TYPE "UDT_Service_ControlBlockMedium"
VERSION : 0.1
   STRUCT
      mode : Int := 1;   //  Service/Mapping selection
      stepOrder { S7_SetPoint := 'False'} : "UDT_Service_StepOrderRawDataMedium";   // Configuration step order
      step { S7_SetPoint := 'False'} : "UDT_Service_StepRawDataMedium" := ([([16#FFFFFFFF], [16#FFFFFFFF], [16#FFFFFFFF], [16#FFFFFFFF]), ([16#FFFFFFFF], [16#FFFFFFFF], [16#FFFFFFFF], [16#FFFFFFFF]), ([16#FFFFFFFF], [16#FFFFFFFF], [16#FFFFFFFF], [16#FFFFFFFF]), ([16#FFFFFFFF], [16#FFFFFFFF], [16#FFFFFFFF], [16#FFFFFFFF]), ([16#FFFFFFFF], [16#FFFFFFFF], [16#FFFFFFFF], [16#FFFFFFFF]), ([16#FFFFFFFF], [16#FFFFFFFF], [16#FFFFFFFF], [16#FFFFFFFF]), ([16#FFFFFFFF], [16#FFFFFFFF], [16#FFFFFFFF], [16#FFFFFFFF]), ([16#FFFFFFFF], [16#FFFFFFFF], [16#FFFFFFFF], [16#FFFFFFFF]), ([16#FFFFFFFF], [16#FFFFFFFF], [16#FFFFFFFF], [16#FFFFFFFF]), ([16#FFFFFFFF], [16#FFFFFFFF], [16#FFFFFFFF], [16#FFFFFFFF]), ([16#FFFFFFFF], [16#FFFFFFFF], [16#FFFFFFFF], [16#FFFFFFFF]), ([16#FFFFFFFF], [16#FFFFFFFF], [16#FFFFFFFF], [16#FFFFFFFF]), ([16#FFFFFFFF], [16#FFFFFFFF], [16#FFFFFFFF], [16#FFFFFFFF]), ([16#FFFFFFFF], [16#FFFFFFFF], [16#FFFFFFFF], [16#FFFFFFFF]), ([16#FFFFFFFF], [16#FFFFFFFF], [16#FFFFFFFF], [16#FFFFFFFF]), ([16#FFFFFFFF], [16#FFFFFFFF], [16#FFFFFFFF], [16#FFFFFFFF]), ([16#FFFFFFFF], [16#FFFFFFFF], [16#FFFFFFFF], [16#FFFFFFFF]), ([16#FFFFFFFF], [16#FFFFFFFF], [16#FFFFFFFF], [16#FFFFFFFF]), ([16#FFFFFFFF], [16#FFFFFFFF], [16#FFFFFFFF], [16#FFFFFFFF]), ([16#FFFFFFFF], [16#FFFFFFFF], [16#FFFFFFFF], [16#FFFFFFFF]), ([16#FFFFFFFF], [16#FFFFFFFF], [16#FFFFFFFF], [16#FFFFFFFF]), ([16#FFFFFFFF], [16#FFFFFFFF], [16#FFFFFFFF], [16#FFFFFFFF]), ([16#FFFFFFFF], [16#FFFFFFFF], [16#FFFFFFFF], [16#FFFFFFFF]), ([16#FFFFFFFF], [16#FFFFFFFF], [16#FFFFFFFF], [16#FFFFFFFF]), ([16#FFFFFFFF], [16#FFFFFFFF], [16#FFFFFFFF], [16#FFFFFFFF]), ([16#FFFFFFFF], [16#FFFFFFFF], [16#FFFFFFFF], [16#FFFFFFFF]), ([16#FFFFFFFF], [16#FFFFFFFF], [16#FFFFFFFF], [16#FFFFFFFF]), ([16#FFFFFFFF], [16#FFFFFFFF], [16#FFFFFFFF], [16#FFFFFFFF]), ([16#FFFFFFFF], [16#FFFFFFFF], [16#FFFFFFFF], [16#FFFFFFFF]), ([16#FFFFFFFF], [16#FFFFFFFF], [16#FFFFFFFF], [16#FFFFFFFF]), ([16#FFFFFFFF], [16#FFFFFFFF], [16#FFFFFFFF], [16#FFFFFFFF]), ([16#FFFFFFFF], [16#FFFFFFFF], [16#FFFFFFFF], [16#FFFFFFFF]), ([16#FFFFFFFF], [16#FFFFFFFF], [16#FFFFFFFF], [16#FFFFFFFF]), ([16#FFFFFFFF], [16#FFFFFFFF], [16#FFFFFFFF], [16#FFFFFFFF]), ([16#FFFFFFFF], [16#FFFFFFFF], [16#FFFFFFFF], [16#FFFFFFFF]), ([16#FFFFFFFF], [16#FFFFFFFF], [16#FFFFFFFF], [16#FFFFFFFF]), ([16#FFFFFFFF], [16#FFFFFFFF], [16#FFFFFFFF], [16#FFFFFFFF]), ([16#FFFFFFFF], [16#FFFFFFFF], [16#FFFFFFFF], [16#FFFFFFFF]), ([16#FFFFFFFF], [16#FFFFFFFF], [16#FFFFFFFF], [16#FFFFFFFF]), ([16#FFFFFFFF], [16#FFFFFFFF], [16#FFFFFFFF], [16#FFFFFFFF]), ([16#FFFFFFFF], [16#FFFFFFFF], [16#FFFFFFFF], [16#FFFFFFFF]), ([16#FFFFFFFF], [16#FFFFFFFF], [16#FFFFFFFF], [16#FFFFFFFF]), ([16#FFFFFFFF], [16#FFFFFFFF], [16#FFFFFFFF], [16#FFFFFFFF]), ([16#FFFFFFFF], [16#FFFFFFFF], [16#FFFFFFFF], [16#FFFFFFFF]), ([16#FFFFFFFF], [16#FFFFFFFF], [16#FFFFFFFF], [16#FFFFFFFF]), ([16#FFFFFFFF], [16#FFFFFFFF], [16#FFFFFFFF], [16#FFFFFFFF]), ([16#FFFFFFFF], [16#FFFFFFFF], [16#FFFFFFFF], [16#FFFFFFFF]), ([16#FFFFFFFF], [16#FFFFFFFF], [16#FFFFFFFF], [16#FFFFFFFF]), ([16#FFFFFFFF], [16#FFFFFFFF], [16#FFFFFFFF], [16#FFFFFFFF]), ([16#FFFFFFFF], [16#FFFFFFFF], [16#FFFFFFFF], [16#FFFFFFFF]), ([16#FFFFFFFF], [16#FFFFFFFF], [16#FFFFFFFF], [16#FFFFFFFF]), ([16#FFFFFFFF], [16#FFFFFFFF], [16#FFFFFFFF], [16#FFFFFFFF]), ([16#FFFFFFFF], [16#FFFFFFFF], [16#FFFFFFFF], [16#FFFFFFFF]), ([16#FFFFFFFF], [16#FFFFFFFF], [16#FFFFFFFF], [16#FFFFFFFF]), ([16#FFFFFFFF], [16#FFFFFFFF], [16#FFFFFFFF], [16#FFFFFFFF]), ([16#FFFFFFFF], [16#FFFFFFFF], [16#FFFFFFFF], [16#FFFFFFFF]), ([16#FFFFFFFF], [16#FFFFFFFF], [16#FFFFFFFF], [16#FFFFFFFF]), ([16#FFFFFFFF], [16#FFFFFFFF], [16#FFFFFFFF], [16#FFFFFFFF]), ([16#FFFFFFFF], [16#FFFFFFFF], [16#FFFFFFFF], [16#FFFFFFFF]), ([16#FFFFFFFF], [16#FFFFFFFF], [16#FFFFFFFF], [16#FFFFFFFF]), ([16#FFFFFFFF], [16#FFFFFFFF], [16#FFFFFFFF], [16#FFFFFFFF]), ([16#FFFFFFFF], [16#FFFFFFFF], [16#FFFFFFFF], [16#FFFFFFFF]), ([16#FFFFFFFF], [16#FFFFFFFF], [16#FFFFFFFF], [16#FFFFFFFF]), ([16#FFFFFFFF], [16#FFFFFFFF], [16#FFFFFFFF], [16#FFFFFFFF]), ([16#FFFFFFFF], [16#FFFFFFFF], [16#FFFFFFFF], [16#FFFFFFFF]), ([16#FFFFFFFF], [16#FFFFFFFF], [16#FFFFFFFF], [16#FFFFFFFF]), ([16#FFFFFFFF], [16#FFFFFFFF], [16#FFFFFFFF], [16#FFFFFFFF]), ([16#FFFFFFFF], [16#FFFFFFFF], [16#FFFFFFFF], [16#FFFFFFFF]), ([16#FFFFFFFF], [16#FFFFFFFF], [16#FFFFFFFF], [16#FFFFFFFF]), ([16#FFFFFFFF], [16#FFFFFFFF], [16#FFFFFFFF], [16#FFFFFFFF]), ([16#FFFFFFFF], [16#FFFFFFFF], [16#FFFFFFFF], [16#FFFFFFFF]), ([16#FFFFFFFF], [16#FFFFFFFF], [16#FFFFFFFF], [16#FFFFFFFF]), ([16#FFFFFFFF], [16#FFFFFFFF], [16#FFFFFFFF], [16#FFFFFFFF]), ([16#FFFFFFFF], [16#FFFFFFFF], [16#FFFFFFFF], [16#FFFFFFFF]), ([16#FFFFFFFF], [16#FFFFFFFF], [16#FFFFFFFF], [16#FFFFFFFF]), ([16#FFFFFFFF], [16#FFFFFFFF], [16#FFFFFFFF], [16#FFFFFFFF]), ([16#FFFFFFFF], [16#FFFFFFFF], [16#FFFFFFFF], [16#FFFFFFFF]), ([16#FFFFFFFF], [16#FFFFFFFF], [16#FFFFFFFF], [16#FFFFFFFF]), ([16#FFFFFFFF], [16#FFFFFFFF], [16#FFFFFFFF], [16#FFFFFFFF]), ([16#FFFFFFFF], [16#FFFFFFFF], [16#FFFFFFFF], [16#FFFFFFFF]), ([16#FFFFFFFF], [16#FFFFFFFF], [16#FFFFFFFF], [16#FFFFFFFF]), ([16#FFFFFFFF], [16#FFFFFFFF], [16#FFFFFFFF], [16#FFFFFFFF]), ([16#FFFFFFFF], [16#FFFFFFFF], [16#FFFFFFFF], [16#FFFFFFFF]), ([16#FFFFFFFF], [16#FFFFFFFF], [16#FFFFFFFF], [16#FFFFFFFF]), ([16#FFFFFFFF], [16#FFFFFFFF], [16#FFFFFFFF], [16#FFFFFFFF]), ([16#FFFFFFFF], [16#FFFFFFFF], [16#FFFFFFFF], [16#FFFFFFFF]), ([16#FFFFFFFF], [16#FFFFFFFF], [16#FFFFFFFF], [16#FFFFFFFF]), ([16#FFFFFFFF], [16#FFFFFFFF], [16#FFFFFFFF], [16#FFFFFFFF]), ([16#FFFFFFFF], [16#FFFFFFFF], [16#FFFFFFFF], [16#FFFFFFFF]), ([16#FFFFFFFF], [16#FFFFFFFF], [16#FFFFFFFF], [16#FFFFFFFF]), ([16#FFFFFFFF], [16#FFFFFFFF], [16#FFFFFFFF], [16#FFFFFFFF]), ([16#FFFFFFFF], [16#FFFFFFFF], [16#FFFFFFFF], [16#FFFFFFFF]), ([16#FFFFFFFF], [16#FFFFFFFF], [16#FFFFFFFF], [16#FFFFFFFF]), ([16#FFFFFFFF], [16#FFFFFFFF], [16#FFFFFFFF], [16#FFFFFFFF]), ([16#FFFFFFFF], [16#FFFFFFFF], [16#FFFFFFFF], [16#FFFFFFFF]), ([16#FFFFFFFF], [16#FFFFFFFF], [16#FFFFFFFF], [16#FFFFFFFF]), ([16#FFFFFFFF], [16#FFFFFFFF], [16#FFFFFFFF], [16#FFFFFFFF]), ([16#FFFFFFFF], [16#FFFFFFFF], [16#FFFFFFFF], [16#FFFFFFFF]), ([16#FFFFFFFF], [16#FFFFFFFF], [16#FFFFFFFF], [16#FFFFFFFF]), ([16#FFFFFFFF], [16#FFFFFFFF], [16#FFFFFFFF], [16#FFFFFFFF])], [((), (), (), ()), ((), (), (), ()), ((), (), (), ()), ((), (), (), ()), ((), (), (), ()), ((), (), (), ()), ((), (), (), ()), ((), (), (), ()), ((), (), (), ()), ((), (), (), ()), ((), (), (), ()), ((), (), (), ()), ((), (), (), ()), ((), (), (), ()), ((), (), (), ()), ((), (), (), ()), ((), (), (), ()), ((), (), (), ()), ((), (), (), ()), ((), (), (), ()), ((), (), (), ()), ((), (), (), ()), ((), (), (), ()), ((), (), (), ()), ((), (), (), ()), ((), (), (), ()), ((), (), (), ()), ((), (), (), ()), ((), (), (), ()), ((), (), (), ()), ((), (), (), ()), ((), (), (), ())]);   // Configuration steps
      procedure { S7_SetPoint := 'False'} : "UDT_Service_ProcedureRawDataMedium";   // Configuration procedures
      configurationParameterData { S7_SetPoint := 'False'} : "UDT_Service_ParameterDataMedium";   // Configuration parameters
      processValueInData { S7_SetPoint := 'False'} : "UDT_Service_ValueDataMedium";   // ProcessIn Values
      processValueOutData { S7_SetPoint := 'False'} : "UDT_Service_ValueDataMedium";   // ProcessOut Values
      reportValueData { S7_SetPoint := 'False'} : "UDT_Service_ValueDataMedium";   // Report Values
      serviceInteraction : Array[1..30] of DWord;   // Service Interaction Information Variable
      plcGuid : String;   // PLC Guid value stored from the tool, used to find the PLC name changes
      serviceGuid : String;   // Service Guid value stored from the tool, used to find the setup DB name changes
      serviceDbNumber : Int;   // Linked Service IDB number stored from the tool, used to find the service name changes
   END_STRUCT;

END_TYPE

